DATA_BLOCK "naut_SfcAltPriority_DB"
{ S7_Optimized_Access := 'TRUE' }
VERSION : 0.1
"naut_SfcAltPriority"

BEGIN

END_DATA_BLOCK
